(*~
	<docu>
		<summary>
			Clears a parameter request.
		</summary>
	</docu>
~*)
FUNCTION TcoAteqG6_ClearParameterRequest_v_3_5_x : BOOL
VAR_IN_OUT
	inoRequest : TcoAteqG6_ParameterRequest_v_3_5_x;
END_VAR
VAR
	i : INT;
END_VAR

inoRequest.Count := 0;
FOR i := 0 TO 34 DO
	inoRequest.Ids[i] := 0;
END_FOR
TcoAteqG6_ClearParameterRequest_v_3_5_x := TRUE;

END_FUNCTION

(* stored: Version 1.1.0.1, ProductVersion 3.1.4024.12
   POU TcoAteqG6_ClearParameterRequest_v_3_5_x: Id {6791b5a3-76d9-47bc-a833-ff921690e5a6}, SpecialFunc None *)
